Fanuc KAREL source: compact_preamble.KL

PROGRAM KX00026
%PRIORITY=20
%NOLOCKGROUP
VAR
I:INTEGER;J:INTEGER;B:BOOLEAN
F : FILE
S : STRING[80]
P : XYZWPR
BEGIN
I=1
END KX00026
